Fanuc KAREL source: KB00039.KL

PROGRAM KB00039
%NOLOCKGROUP
%ENVIRONMENT STRNG
VAR
  P1: STRING[80]
  P2: CONFIG
  P3: INTEGER
BEGIN
  P1 = 'A'
  P3 = 1
  CNV_STR_CONF(P1, P2, P3)
END KB00039
